(* IEC 61131-3 sources: codesys-ai-industrial-robot-control/plc/src, 6 files *)

(* ---- ST_Recipe_Cell.st ---- *)
TYPE ST_Recipe_Cell :
STRUCT
    lrBeltSpeed : LREAL; // GVL_Params.lrBeltSpeed
    lrApproachHeight : LREAL; // GVL_Params.lrApproachHeight
    lrPickDepth : LREAL; // GVL_Params.lrPickDepth
    lrLinVelocity : LREAL; // GVL_Params.lrLinVelocity
    lrLinAccel : LREAL; // GVL_Params.lrLinAccel
    lrLinJerk : LREAL; // GVL_Params.lrLinJerk
    lrPtpVelFactor : LREAL; // GVL_Params.lrPtpVelFactor
    rConfidenceThreshold : REAL; // GVL_Params.rConfidenceThreshold
    tDecisionDeadline : TIME; // GVL_Params.tDecisionDeadline
    tVacuumTimeout : TIME; // GVL_Params.tVacuumTimeout
    lrFollowErrWarn : LREAL; // GVL_Params.lrFollowErrWarn
    lrFollowErrFault : LREAL; // GVL_Params.lrFollowErrFault
    tFeedbackTimeout : TIME; // GVL_Params.tFeedbackTimeout
END_STRUCT
END_TYPE

(* ---- GVL_Recipe_Cell.st ---- *)
// Recipes 'Cell', generated by codesys-mcp-toolkit (create_recipes). RETAIN: values saved from the HMI survive a power cycle.
VAR_GLOBAL RETAIN
    aRecipes : ARRAY[0..1] OF ST_Recipe_Cell := [(lrBeltSpeed := 100.0, lrApproachHeight := 80.0, lrPickDepth := 5.0, lrLinVelocity := 500.0, lrLinAccel := 2000.0, lrLinJerk := 20000.0, lrPtpVelFactor := 0.5, rConfidenceThreshold := 0.6, tDecisionDeadline := T#2S500MS, tVacuumTimeout := T#500MS, lrFollowErrWarn := 2.0, lrFollowErrFault := 5.0, tFeedbackTimeout := T#500MS), (lrBeltSpeed := 200.0, lrApproachHeight := 80.0, lrPickDepth := 5.0, lrLinVelocity := 800.0, lrLinAccel := 3000.0, lrLinJerk := 20000.0, lrPtpVelFactor := 0.8, rConfidenceThreshold := 0.6, tDecisionDeadline := T#2S500MS, tVacuumTimeout := T#500MS, lrFollowErrWarn := 2.0, lrFollowErrFault := 5.0, tFeedbackTimeout := T#500MS)];
END_VAR
VAR_GLOBAL CONSTANT
    asNames : ARRAY[0..1] OF STRING(32) := ['Standard', 'HighSpeed'];
    iCount : INT := 2;
END_VAR

(* ---- PRG_HMI_Alarms.st ---- *)
PROGRAM PRG_HMI_Alarms
// Generated by codesys-mcp-toolkit for the HMI screen 'Alarms' (42 variables). Rebuilt on every export.
VAR
    iMachine : INT; // the machine's state: 0 idle, 1.. the states in order
    sV1 : STRING(80); // GVL_HmiView.sState
    sV2 : STRING(80); // GVL_HmiView.sMode
    rV3 : REAL; // GVL_HmiView.sNewestAlarm
END_VAR

IF GVL_HmiView.xAborted THEN iMachine := 1; ELSIF GVL_HmiView.xHeld THEN iMachine := 2; ELSIF GVL_HmiView.xActing THEN iMachine := 3; ELSIF GVL_HmiView.xManual THEN iMachine := 4; ELSIF GVL_HmiView.xExecute THEN iMachine := 5; ELSIF GVL_HmiView.xIdle THEN iMachine := 6; ELSE iMachine := 0; END_IF
sV1 := TO_STRING(GVL_HmiView.sState);
sV2 := TO_STRING(GVL_HmiView.sMode);
rV3 := ANY_TO_REAL(GVL_HmiView.sNewestAlarm);

(* ---- PRG_HMI_Overview.st ---- *)
PROGRAM PRG_HMI_Overview
// Generated by codesys-mcp-toolkit for the HMI screen 'Overview' (49 variables). Rebuilt on every export.
VAR
    iMachine : INT; // the machine's state: 0 idle, 1.. the states in order
    sV1 : STRING(80); // GVL_HmiView.sState
    sV2 : STRING(80); // GVL_HmiView.sMode
    rV3 : REAL; // GVL_HmiView.uiPlaced
    rV4 : REAL; // GVL_Bridge.lrBeltVel
    rV5 : REAL; // GVL_HmiView.uiPlaced
    rV6 : REAL; // GVL_Bridge.lrBeltVel
    iP7 : INT; // GVL_Bridge.lrBeltVel
    rV8 : REAL; // GVL_HmiView.uiPlaced
    rV9 : REAL; // PRG_Main.fbCell.aBins[0].uiCount
    xB10 : BOOL; // PRG_Main.fbCell.aBins[0].uiCount >= 27
    iP11 : INT; // PRG_Main.fbCell.aBins[0].uiCount
    xB12 : BOOL; // PRG_Main.fbCell.aBins[0].uiCount >= 27
    rV13 : REAL; // PRG_Main.fbCell.aBins[1].uiCount
    xB14 : BOOL; // PRG_Main.fbCell.aBins[1].uiCount >= 27
    iP15 : INT; // PRG_Main.fbCell.aBins[1].uiCount
    xB16 : BOOL; // PRG_Main.fbCell.aBins[1].uiCount >= 27
    rV17 : REAL; // PRG_Main.fbCell.aBins[2].uiCount
    xB18 : BOOL; // PRG_Main.fbCell.aBins[2].uiCount >= 27
    iP19 : INT; // PRG_Main.fbCell.aBins[2].uiCount
    xB20 : BOOL; // PRG_Main.fbCell.aBins[2].uiCount >= 27
    rV21 : REAL; // PRG_Main.fbCell.aBins[3].uiCount
    xB22 : BOOL; // PRG_Main.fbCell.aBins[3].uiCount >= 27
    iP23 : INT; // PRG_Main.fbCell.aBins[3].uiCount
    xB24 : BOOL; // PRG_Main.fbCell.aBins[3].uiCount >= 27
    rV25 : REAL; // PRG_Main.fbCell.aBins[4].uiCount
    xB26 : BOOL; // PRG_Main.fbCell.aBins[4].uiCount >= 27
    iP27 : INT; // PRG_Main.fbCell.aBins[4].uiCount
    xB28 : BOOL; // PRG_Main.fbCell.aBins[4].uiCount >= 27
    rV29 : REAL; // PRG_Main.fbCell.aBins[5].uiCount
    xB30 : BOOL; // PRG_Main.fbCell.aBins[5].uiCount >= 27
    iP31 : INT; // PRG_Main.fbCell.aBins[5].uiCount
    xB32 : BOOL; // PRG_Main.fbCell.aBins[5].uiCount >= 27
END_VAR

IF GVL_HmiView.xAborted THEN iMachine := 1; ELSIF GVL_HmiView.xHeld THEN iMachine := 2; ELSIF GVL_HmiView.xActing THEN iMachine := 3; ELSIF GVL_HmiView.xManual THEN iMachine := 4; ELSIF GVL_HmiView.xExecute THEN iMachine := 5; ELSIF GVL_HmiView.xIdle THEN iMachine := 6; ELSE iMachine := 0; END_IF
sV1 := TO_STRING(GVL_HmiView.sState);
sV2 := TO_STRING(GVL_HmiView.sMode);
rV3 := ANY_TO_REAL(GVL_HmiView.uiPlaced);
rV4 := ANY_TO_REAL(GVL_Bridge.lrBeltVel);
rV5 := ANY_TO_REAL(GVL_HmiView.uiPlaced);
rV6 := ANY_TO_REAL(GVL_Bridge.lrBeltVel);
iP7 := REAL_TO_INT(LIMIT(0.0, (ANY_TO_REAL(GVL_Bridge.lrBeltVel) - (0.0)) / (150.0), 1.0) * 374.0);
rV8 := ANY_TO_REAL(GVL_HmiView.uiPlaced);
rV9 := ANY_TO_REAL(PRG_Main.fbCell.aBins[0].uiCount);
xB10 := ANY_TO_REAL(PRG_Main.fbCell.aBins[0].uiCount) >= 27.0;
iP11 := REAL_TO_INT(LIMIT(0.0, (ANY_TO_REAL(PRG_Main.fbCell.aBins[0].uiCount) - (0.0)) / (30.0), 1.0) * 80.0);
xB12 := ANY_TO_REAL(PRG_Main.fbCell.aBins[0].uiCount) >= 27.0;
rV13 := ANY_TO_REAL(PRG_Main.fbCell.aBins[1].uiCount);
xB14 := ANY_TO_REAL(PRG_Main.fbCell.aBins[1].uiCount) >= 27.0;
iP15 := REAL_TO_INT(LIMIT(0.0, (ANY_TO_REAL(PRG_Main.fbCell.aBins[1].uiCount) - (0.0)) / (30.0), 1.0) * 80.0);
xB16 := ANY_TO_REAL(PRG_Main.fbCell.aBins[1].uiCount) >= 27.0;
rV17 := ANY_TO_REAL(PRG_Main.fbCell.aBins[2].uiCount);
xB18 := ANY_TO_REAL(PRG_Main.fbCell.aBins[2].uiCount) >= 27.0;
iP19 := REAL_TO_INT(LIMIT(0.0, (ANY_TO_REAL(PRG_Main.fbCell.aBins[2].uiCount) - (0.0)) / (30.0), 1.0) * 80.0);
xB20 := ANY_TO_REAL(PRG_Main.fbCell.aBins[2].uiCount) >= 27.0;
rV21 := ANY_TO_REAL(PRG_Main.fbCell.aBins[3].uiCount);
xB22 := ANY_TO_REAL(PRG_Main.fbCell.aBins[3].uiCount) >= 27.0;
iP23 := REAL_TO_INT(LIMIT(0.0, (ANY_TO_REAL(PRG_Main.fbCell.aBins[3].uiCount) - (0.0)) / (30.0), 1.0) * 80.0);
xB24 := ANY_TO_REAL(PRG_Main.fbCell.aBins[3].uiCount) >= 27.0;
rV25 := ANY_TO_REAL(PRG_Main.fbCell.aBins[4].uiCount);
xB26 := ANY_TO_REAL(PRG_Main.fbCell.aBins[4].uiCount) >= 27.0;
iP27 := REAL_TO_INT(LIMIT(0.0, (ANY_TO_REAL(PRG_Main.fbCell.aBins[4].uiCount) - (0.0)) / (30.0), 1.0) * 80.0);
xB28 := ANY_TO_REAL(PRG_Main.fbCell.aBins[4].uiCount) >= 27.0;
rV29 := ANY_TO_REAL(PRG_Main.fbCell.aBins[5].uiCount);
xB30 := ANY_TO_REAL(PRG_Main.fbCell.aBins[5].uiCount) >= 27.0;
iP31 := REAL_TO_INT(LIMIT(0.0, (ANY_TO_REAL(PRG_Main.fbCell.aBins[5].uiCount) - (0.0)) / (30.0), 1.0) * 80.0);
xB32 := ANY_TO_REAL(PRG_Main.fbCell.aBins[5].uiCount) >= 27.0;

(* ---- PRG_HMI_Robot.st ---- *)
PROGRAM PRG_HMI_Robot
// Generated by codesys-mcp-toolkit for the HMI screen 'Robot' (49 variables). Rebuilt on every export.
VAR
    iMachine : INT; // the machine's state: 0 idle, 1.. the states in order
    sV1 : STRING(80); // GVL_HmiView.sState
    sV2 : STRING(80); // GVL_HmiView.sMode
    rV3 : REAL; // GVL_HmiView.uiPlaced
    rV4 : REAL; // GVL_Bridge.aJointPosSp[1]
    iP5 : INT; // GVL_Bridge.aJointPosSp[1]
    rV6 : REAL; // GVL_Bridge.aJointPosSp[2]
    iP7 : INT; // GVL_Bridge.aJointPosSp[2]
    rV8 : REAL; // GVL_Bridge.aJointPosSp[3]
    iP9 : INT; // GVL_Bridge.aJointPosSp[3]
    rV10 : REAL; // GVL_Bridge.aJointPosSp[4]
    iP11 : INT; // GVL_Bridge.aJointPosSp[4]
    rV12 : REAL; // GVL_Bridge.aJointPosSp[5]
    iP13 : INT; // GVL_Bridge.aJointPosSp[5]
    rV14 : REAL; // GVL_Bridge.aJointPosSp[6]
    iP15 : INT; // GVL_Bridge.aJointPosSp[6]
    rV16 : REAL; // GVL_Bridge.aFollowingError[1]
    xB17 : BOOL; // GVL_Bridge.aFollowingError[1] >= 2
    iP18 : INT; // GVL_Bridge.aFollowingError[1]
    xB19 : BOOL; // GVL_Bridge.aFollowingError[1] >= 2
    rV20 : REAL; // GVL_Bridge.aFollowingError[2]
    xB21 : BOOL; // GVL_Bridge.aFollowingError[2] >= 2
    iP22 : INT; // GVL_Bridge.aFollowingError[2]
    xB23 : BOOL; // GVL_Bridge.aFollowingError[2] >= 2
    rV24 : REAL; // GVL_Bridge.aFollowingError[3]
    xB25 : BOOL; // GVL_Bridge.aFollowingError[3] >= 2
    iP26 : INT; // GVL_Bridge.aFollowingError[3]
    xB27 : BOOL; // GVL_Bridge.aFollowingError[3] >= 2
    rV28 : REAL; // GVL_Bridge.aFollowingError[4]
    xB29 : BOOL; // GVL_Bridge.aFollowingError[4] >= 2
    iP30 : INT; // GVL_Bridge.aFollowingError[4]
    xB31 : BOOL; // GVL_Bridge.aFollowingError[4] >= 2
    rV32 : REAL; // GVL_Bridge.aFollowingError[5]
    xB33 : BOOL; // GVL_Bridge.aFollowingError[5] >= 2
    iP34 : INT; // GVL_Bridge.aFollowingError[5]
    xB35 : BOOL; // GVL_Bridge.aFollowingError[5] >= 2
    rV36 : REAL; // GVL_Bridge.aFollowingError[6]
    xB37 : BOOL; // GVL_Bridge.aFollowingError[6] >= 2
    iP38 : INT; // GVL_Bridge.aFollowingError[6]
    xB39 : BOOL; // GVL_Bridge.aFollowingError[6] >= 2
    rV40 : REAL; // GVL_Hmi.rOverride
    rV41 : REAL; // GVL_Bridge.iWorstJoint
    rV42 : REAL; // GVL_Bridge.stVision.usiClass
    rV43 : REAL; // GVL_Bridge.stVision.rConfidence
    rV44 : REAL; // GVL_Bridge.stVision.lrX
END_VAR

IF GVL_HmiView.xAborted THEN iMachine := 1; ELSIF GVL_HmiView.xHeld THEN iMachine := 2; ELSIF GVL_HmiView.xActing THEN iMachine := 3; ELSIF GVL_HmiView.xManual THEN iMachine := 4; ELSIF GVL_HmiView.xExecute THEN iMachine := 5; ELSIF GVL_HmiView.xIdle THEN iMachine := 6; ELSE iMachine := 0; END_IF
sV1 := TO_STRING(GVL_HmiView.sState);
sV2 := TO_STRING(GVL_HmiView.sMode);
rV3 := ANY_TO_REAL(GVL_HmiView.uiPlaced);
rV4 := ANY_TO_REAL(GVL_Bridge.aJointPosSp[1]);
iP5 := REAL_TO_INT(LIMIT(0.0, (ANY_TO_REAL(GVL_Bridge.aJointPosSp[1]) - (-180.0)) / (360.0), 1.0) * 80.0);
rV6 := ANY_TO_REAL(GVL_Bridge.aJointPosSp[2]);
iP7 := REAL_TO_INT(LIMIT(0.0, (ANY_TO_REAL(GVL_Bridge.aJointPosSp[2]) - (-180.0)) / (360.0), 1.0) * 80.0);
rV8 := ANY_TO_REAL(GVL_Bridge.aJointPosSp[3]);
iP9 := REAL_TO_INT(LIMIT(0.0, (ANY_TO_REAL(GVL_Bridge.aJointPosSp[3]) - (-180.0)) / (360.0), 1.0) * 80.0);
rV10 := ANY_TO_REAL(GVL_Bridge.aJointPosSp[4]);
iP11 := REAL_TO_INT(LIMIT(0.0, (ANY_TO_REAL(GVL_Bridge.aJointPosSp[4]) - (-360.0)) / (720.0), 1.0) * 80.0);
rV12 := ANY_TO_REAL(GVL_Bridge.aJointPosSp[5]);
iP13 := REAL_TO_INT(LIMIT(0.0, (ANY_TO_REAL(GVL_Bridge.aJointPosSp[5]) - (-180.0)) / (360.0), 1.0) * 80.0);
rV14 := ANY_TO_REAL(GVL_Bridge.aJointPosSp[6]);
iP15 := REAL_TO_INT(LIMIT(0.0, (ANY_TO_REAL(GVL_Bridge.aJointPosSp[6]) - (-360.0)) / (720.0), 1.0) * 80.0);
rV16 := ANY_TO_REAL(GVL_Bridge.aFollowingError[1]);
xB17 := ANY_TO_REAL(GVL_Bridge.aFollowingError[1]) >= 2.0;
iP18 := REAL_TO_INT(LIMIT(0.0, (ANY_TO_REAL(GVL_Bridge.aFollowingError[1]) - (0.0)) / (6.0), 1.0) * 80.0);
xB19 := ANY_TO_REAL(GVL_Bridge.aFollowingError[1]) >= 2.0;
rV20 := ANY_TO_REAL(GVL_Bridge.aFollowingError[2]);
xB21 := ANY_TO_REAL(GVL_Bridge.aFollowingError[2]) >= 2.0;
iP22 := REAL_TO_INT(LIMIT(0.0, (ANY_TO_REAL(GVL_Bridge.aFollowingError[2]) - (0.0)) / (6.0), 1.0) * 80.0);
xB23 := ANY_TO_REAL(GVL_Bridge.aFollowingError[2]) >= 2.0;
rV24 := ANY_TO_REAL(GVL_Bridge.aFollowingError[3]);
xB25 := ANY_TO_REAL(GVL_Bridge.aFollowingError[3]) >= 2.0;
iP26 := REAL_TO_INT(LIMIT(0.0, (ANY_TO_REAL(GVL_Bridge.aFollowingError[3]) - (0.0)) / (6.0), 1.0) * 80.0);
xB27 := ANY_TO_REAL(GVL_Bridge.aFollowingError[3]) >= 2.0;
rV28 := ANY_TO_REAL(GVL_Bridge.aFollowingError[4]);
xB29 := ANY_TO_REAL(GVL_Bridge.aFollowingError[4]) >= 2.0;
iP30 := REAL_TO_INT(LIMIT(0.0, (ANY_TO_REAL(GVL_Bridge.aFollowingError[4]) - (0.0)) / (6.0), 1.0) * 80.0);
xB31 := ANY_TO_REAL(GVL_Bridge.aFollowingError[4]) >= 2.0;
rV32 := ANY_TO_REAL(GVL_Bridge.aFollowingError[5]);
xB33 := ANY_TO_REAL(GVL_Bridge.aFollowingError[5]) >= 2.0;
iP34 := REAL_TO_INT(LIMIT(0.0, (ANY_TO_REAL(GVL_Bridge.aFollowingError[5]) - (0.0)) / (6.0), 1.0) * 80.0);
xB35 := ANY_TO_REAL(GVL_Bridge.aFollowingError[5]) >= 2.0;
rV36 := ANY_TO_REAL(GVL_Bridge.aFollowingError[6]);
xB37 := ANY_TO_REAL(GVL_Bridge.aFollowingError[6]) >= 2.0;
iP38 := REAL_TO_INT(LIMIT(0.0, (ANY_TO_REAL(GVL_Bridge.aFollowingError[6]) - (0.0)) / (6.0), 1.0) * 80.0);
xB39 := ANY_TO_REAL(GVL_Bridge.aFollowingError[6]) >= 2.0;
rV40 := ANY_TO_REAL(GVL_Hmi.rOverride);
rV41 := ANY_TO_REAL(GVL_Bridge.iWorstJoint);
rV42 := ANY_TO_REAL(GVL_Bridge.stVision.usiClass);
rV43 := ANY_TO_REAL(GVL_Bridge.stVision.rConfidence);
rV44 := ANY_TO_REAL(GVL_Bridge.stVision.lrX);

(* ---- PRG_Recipe_Cell.st ---- *)
PROGRAM PRG_Recipe_Cell
// Set iApply to a recipe's index to write it to the variables; set iSave to store the variables in it.
VAR
    iApply : INT := -1;
    iSave : INT := -1;
    iActive : INT := -1; // the recipe applied last
    sActive : STRING(32);
    p0 : POINTER TO LREAL; // GVL_Params.lrBeltSpeed
    p1 : POINTER TO LREAL; // GVL_Params.lrApproachHeight
    p2 : POINTER TO LREAL; // GVL_Params.lrPickDepth
    p3 : POINTER TO LREAL; // GVL_Params.lrLinVelocity
    p4 : POINTER TO LREAL; // GVL_Params.lrLinAccel
    p5 : POINTER TO LREAL; // GVL_Params.lrLinJerk
    p6 : POINTER TO LREAL; // GVL_Params.lrPtpVelFactor
    p7 : POINTER TO REAL; // GVL_Params.rConfidenceThreshold
    p8 : POINTER TO TIME; // GVL_Params.tDecisionDeadline
    p9 : POINTER TO TIME; // GVL_Params.tVacuumTimeout
    p10 : POINTER TO LREAL; // GVL_Params.lrFollowErrWarn
    p11 : POINTER TO LREAL; // GVL_Params.lrFollowErrFault
    p12 : POINTER TO TIME; // GVL_Params.tFeedbackTimeout
END_VAR

p0 := ADR(GVL_Params.lrBeltSpeed);
p1 := ADR(GVL_Params.lrApproachHeight);
p2 := ADR(GVL_Params.lrPickDepth);
p3 := ADR(GVL_Params.lrLinVelocity);
p4 := ADR(GVL_Params.lrLinAccel);
p5 := ADR(GVL_Params.lrLinJerk);
p6 := ADR(GVL_Params.lrPtpVelFactor);
p7 := ADR(GVL_Params.rConfidenceThreshold);
p8 := ADR(GVL_Params.tDecisionDeadline);
p9 := ADR(GVL_Params.tVacuumTimeout);
p10 := ADR(GVL_Params.lrFollowErrWarn);
p11 := ADR(GVL_Params.lrFollowErrFault);
p12 := ADR(GVL_Params.tFeedbackTimeout);
IF iApply >= 0 AND iApply < 2 THEN
    p0^ := GVL_Recipe_Cell.aRecipes[iApply].lrBeltSpeed;
    p1^ := GVL_Recipe_Cell.aRecipes[iApply].lrApproachHeight;
    p2^ := GVL_Recipe_Cell.aRecipes[iApply].lrPickDepth;
    p3^ := GVL_Recipe_Cell.aRecipes[iApply].lrLinVelocity;
    p4^ := GVL_Recipe_Cell.aRecipes[iApply].lrLinAccel;
    p5^ := GVL_Recipe_Cell.aRecipes[iApply].lrLinJerk;
    p6^ := GVL_Recipe_Cell.aRecipes[iApply].lrPtpVelFactor;
    p7^ := GVL_Recipe_Cell.aRecipes[iApply].rConfidenceThreshold;
    p8^ := GVL_Recipe_Cell.aRecipes[iApply].tDecisionDeadline;
    p9^ := GVL_Recipe_Cell.aRecipes[iApply].tVacuumTimeout;
    p10^ := GVL_Recipe_Cell.aRecipes[iApply].lrFollowErrWarn;
    p11^ := GVL_Recipe_Cell.aRecipes[iApply].lrFollowErrFault;
    p12^ := GVL_Recipe_Cell.aRecipes[iApply].tFeedbackTimeout;
    iActive := iApply;
    sActive := GVL_Recipe_Cell.asNames[iApply];
END_IF
iApply := -1;
IF iSave >= 0 AND iSave < 2 THEN
    GVL_Recipe_Cell.aRecipes[iSave].lrBeltSpeed := p0^;
    GVL_Recipe_Cell.aRecipes[iSave].lrApproachHeight := p1^;
    GVL_Recipe_Cell.aRecipes[iSave].lrPickDepth := p2^;
    GVL_Recipe_Cell.aRecipes[iSave].lrLinVelocity := p3^;
    GVL_Recipe_Cell.aRecipes[iSave].lrLinAccel := p4^;
    GVL_Recipe_Cell.aRecipes[iSave].lrLinJerk := p5^;
    GVL_Recipe_Cell.aRecipes[iSave].lrPtpVelFactor := p6^;
    GVL_Recipe_Cell.aRecipes[iSave].rConfidenceThreshold := p7^;
    GVL_Recipe_Cell.aRecipes[iSave].tDecisionDeadline := p8^;
    GVL_Recipe_Cell.aRecipes[iSave].tVacuumTimeout := p9^;
    GVL_Recipe_Cell.aRecipes[iSave].lrFollowErrWarn := p10^;
    GVL_Recipe_Cell.aRecipes[iSave].lrFollowErrFault := p11^;
    GVL_Recipe_Cell.aRecipes[iSave].tFeedbackTimeout := p12^;
END_IF
iSave := -1;
